(*
SPDX-FileCopyrightText: c 2026 Oleksandr Tiutyk <trofimich@gmail.com>
SPDX-License-Identifier: MIT
License: https://opensource.org/license/mit
*)

(*!
<summary>Checks raw membership without changing LIFO order.</summary>
<description>
Borrows a group-owned stack reserved for this case. Use from one task at a stable address.
Teardown clears the stack and test-owned resources before publication.
</description>
*)

{attribute 'no_assign'}
{attribute 'no_explicit_call' := 'do not call this function block directly'}
FUNCTION_BLOCK StackContainsTest EXTENDS TOF_Testing.SingleCycleTest
VAR_STAT
	{attribute 'hide'}
	_ClassName : STRING := __POUNAME();
END_VAR
VAR
	_Stack : TOF_Collections.IStack;
END_VAR

(*!
<summary>Clears the fixture before the runner publishes the result.</summary>
<description>
Also runs after an unexpected exception interrupts the case.
</description>
*)
METHOD PROTECTED AfterTest
_Stack.Clear();
END_METHOD

//! <summary>Borrows the concrete class name. Callers must not modify it.</summary>
{attribute 'monitoring' := 'call'}
PROPERTY ClassName : REFERENCE TO STRING
GET
ClassName REF= _ClassName;
END_GET
END_PROPERTY

(*!
<summary>Checks raw membership without changing LIFO order.</summary>
*)
METHOD PROTECTED ExecuteTest
VAR
	values : ARRAY [1..4] OF INT := [11, 22, 33, 44];
END_VAR
Assert.ThatBool(
	actual := _Stack.Contains(value := values[1]),
	message := "An empty stack must report absence"
).IsFalse();

_Stack.PushCopy(value := values[1]);
_Stack.PushCopy(value := values[2]);
_Stack.PushCopy(value := values[3]);

Assert.ThatBool(
	actual := _Stack.Contains(value := values[1]),
	message := "Contains must find the bottom value"
).IsTrue();

Assert.ThatBool(
	actual := _Stack.Contains(value := values[3]),
	message := "Contains must find the top value"
).IsTrue();

Assert.ThatBool(
	actual := _Stack.Contains(value := values[4]),
	message := "Contains must reject an absent value"
).IsFalse();

Assert.ThatDInt(
	actual := _Stack.Length,
	message := "Lookup must preserve all three entries"
).ToBe(expected := DINT#3);
END_METHOD

(*!
<summary>Binds the stack fixture for this case.</summary>
<description>
Stores a borrowed interface without invoking the fixture. The owning group keeps it alive and
reserves it for this case. TestElement initializes the name and parent.
</description>
<param name="name">Display name of this case.</param>
<param name="parent">Group that owns this case.</param>
<param name="stack">Required live stack reserved for this case.</param>
*)
METHOD FB_init : BOOL
VAR_INPUT
	bInitRetains: BOOL; // TRUE: the retain variables are initialized (reset warm / reset cold)
	bInCopyCode: BOOL; // TRUE: the instance will be copied to the copy code afterward (online change)
	name : WSTRING;
	parent : TOF_Testing.ITestElement;
	stack : TOF_Collections.IStack;
END_VAR
_Stack := stack;
FB_init := TRUE;
END_METHOD

//! <summary>Borrows the compiler-initialized namespace name. Callers must not modify it.</summary>
{attribute 'monitoring' := 'call'}
PROPERTY NamespaceName : REFERENCE TO STRING
GET
NamespaceName REF= CurrentNamespace.Name;
END_GET
END_PROPERTY

//! <summary>Reports the concrete instance size in bytes.</summary>
{attribute 'monitoring' := 'call'}
PROPERTY SelfSize : ULINT
GET
SelfSize := XSIZEOF(THIS^);
END_GET
END_PROPERTY

END_FUNCTION_BLOCK

(* stored: Version 1.1.0.1, ProductVersion 3.1.4026.21
   POU StackContainsTest: Id {80e60297-9d78-4565-8d32-876b091a8528}, SpecialFunc None
   Method AfterTest: Id {641a6d8e-f8ad-453f-a92f-8bf85785b590}
   Property ClassName: Id {3701ee6a-5b6f-4245-a2c3-02b143b51988}
   Get Get: Id {0cc70852-ef34-47a4-ad43-3a207a287e87}
   Method ExecuteTest: Id {5302e7c1-15e5-4c2b-98c8-c5cbdd9a547d}
   Method FB_init: Id {3b596234-5fbf-4a79-bab8-49688380f6c0}
   Property NamespaceName: Id {7661b4a4-b296-42fd-9426-1f70450980e7}
   Get Get: Id {c87ff028-cd82-4ab9-adc3-019b85856239}
   Property SelfSize: Id {1224eca4-50ac-4146-a465-8d4b0d2023d9}
   Get Get: Id {dc9ed70d-1e23-4438-89c8-f1a7728e2ca2} *)
